Fanuc KAREL source: KD00033.KL

PROGRAM KD00033
%NOLOCKGROUP
VAR
  I: INTEGER
  J: INTEGER
  B: BOOLEAN
  R: REAL
  S: STRING[80]
BEGIN
  CONDITION[1]:
  WHEN DIN[1] = ON DO
    I = 1
  ENDCONDITION
END KD00033
